(* IEC 61131-3 sources: plcassist-cli/packages/volt-lsp-iec/test-corpus/pro2193/Device/Plc Logic/Application/09 Misc/Library Manager/Standard64, 25 files *)

(* ---- ATOMICREADLINT.fun ---- *)
FUNCTION ATOMICREADLINT : LINT
VAR_INPUT
	PSRC : POINTER TO LINT;
END_VAR
END_FUNCTION

(* ---- ATOMICREADLREAL.fun ---- *)
FUNCTION ATOMICREADLREAL : LREAL
VAR_INPUT
	PSRC : POINTER TO LREAL;
END_VAR
END_FUNCTION

(* ---- ATOMICREADLTIME.fun ---- *)
FUNCTION ATOMICREADLTIME : LTIME
VAR_INPUT
	PSRC : POINTER TO LTIME;
END_VAR
END_FUNCTION

(* ---- ATOMICREADLWORD.fun ---- *)
FUNCTION ATOMICREADLWORD : LWORD
VAR_INPUT
	PSRC : POINTER TO LWORD;
END_VAR
END_FUNCTION

(* ---- ATOMICREADULINT.fun ---- *)
FUNCTION ATOMICREADULINT : ULINT
VAR_INPUT
	PSRC : POINTER TO ULINT;
END_VAR
END_FUNCTION

(* ---- ATOMICWRITELINT.fun ---- *)
FUNCTION ATOMICWRITELINT : BOOL
VAR_INPUT
	PDEST : POINTER TO LINT;
	LIVALUE : LINT;
END_VAR
END_FUNCTION

(* ---- ATOMICWRITELREAL.fun ---- *)
FUNCTION ATOMICWRITELREAL : BOOL
VAR_INPUT
	PDEST : POINTER TO LREAL;
	LRVALUE : LREAL;
END_VAR
END_FUNCTION

(* ---- ATOMICWRITELTIME.fun ---- *)
FUNCTION ATOMICWRITELTIME : BOOL
VAR_INPUT
	PDEST : POINTER TO LTIME;
	LTVALUE : LTIME;
END_VAR
END_FUNCTION

(* ---- ATOMICWRITELWORD.fun ---- *)
FUNCTION ATOMICWRITELWORD : BOOL
VAR_INPUT
	PDEST : POINTER TO LWORD;
	LWVALUE : LWORD;
END_VAR
END_FUNCTION

(* ---- ATOMICWRITEULINT.fun ---- *)
FUNCTION ATOMICWRITEULINT : BOOL
VAR_INPUT
	PDEST : POINTER TO ULINT;
	ULIVALUE : ULINT;
END_VAR
END_FUNCTION

(* ---- WCONCAT.fun ---- *)
FUNCTION WCONCAT : WSTRING(255)
VAR_INPUT
	STR1 : WSTRING(255);
	STR2 : WSTRING(255);
END_VAR
END_FUNCTION

(* ---- WDELETE.fun ---- *)
FUNCTION WDELETE : WSTRING(255)
VAR_INPUT
	STR : WSTRING(255);
	LEN : INT;
	POS : INT;
END_VAR
END_FUNCTION

(* ---- WFIND.fun ---- *)
FUNCTION WFIND : INT
VAR_INPUT
	STR1 : WSTRING(255);
	STR2 : WSTRING(255);
END_VAR
END_FUNCTION

(* ---- WINSERT.fun ---- *)
FUNCTION WINSERT : WSTRING(255)
VAR_INPUT
	STR1 : WSTRING(255);
	STR2 : WSTRING(255);
	POS : INT;
END_VAR
END_FUNCTION

(* ---- WLEFT.fun ---- *)
FUNCTION WLEFT : WSTRING(255)
VAR_INPUT
	STR : WSTRING(255);
	SIZE : INT;
END_VAR
END_FUNCTION

(* ---- WLEN.fun ---- *)
FUNCTION WLEN : INT
VAR_INPUT
	STR : WSTRING(255);
END_VAR
END_FUNCTION

(* ---- WMID.fun ---- *)
FUNCTION WMID : WSTRING(255)
VAR_INPUT
	STR : WSTRING(255);
	LEN : INT;
	POS : INT;
END_VAR
END_FUNCTION

(* ---- WREPLACE.fun ---- *)
FUNCTION WREPLACE : WSTRING(255)
VAR_INPUT
	STR1 : WSTRING(255);
	STR2 : WSTRING(255);
	L : INT;
	P : INT;
END_VAR
END_FUNCTION

(* ---- WRIGHT.fun ---- *)
FUNCTION WRIGHT : WSTRING(255)
VAR_INPUT
	STR : WSTRING(255);
	SIZE : INT;
END_VAR
END_FUNCTION

(* ---- LCTD.fb ---- *)
FUNCTION_BLOCK LCTD
VAR_INPUT
	CD : BOOL;
	LOAD : BOOL;
	PV : LWORD;
END_VAR
VAR_OUTPUT
	Q : BOOL;
	CV : LWORD;
END_VAR
VAR
	M : BOOL;
END_VAR
END_FUNCTION_BLOCK

(* ---- LCTU.fb ---- *)
FUNCTION_BLOCK LCTU
VAR_INPUT
	CU : BOOL;
	RESET : BOOL;
	PV : LWORD;
END_VAR
VAR_OUTPUT
	Q : BOOL;
	CV : LWORD;
END_VAR
VAR
	M : BOOL;
END_VAR
END_FUNCTION_BLOCK

(* ---- LCTUD.fb ---- *)
FUNCTION_BLOCK LCTUD
VAR_INPUT
	CU : BOOL;
	CD : BOOL;
	RESET : BOOL;
	LOAD : BOOL;
	PV : LWORD;
END_VAR
VAR_OUTPUT
	QU : BOOL;
	QD : BOOL;
	CV : LWORD;
END_VAR
VAR
	MU : BOOL;
	MD : BOOL;
	RU : BOOL;
	RD : BOOL;
END_VAR
END_FUNCTION_BLOCK

(* ---- LTOF.fb ---- *)
FUNCTION_BLOCK LTOF
VAR_INPUT
	IN : BOOL;
	PT : LTIME;
END_VAR
VAR_OUTPUT
	Q : BOOL;
	ET : LTIME;
END_VAR
VAR
	M : BOOL;
	STARTTIME : LTIME;
END_VAR
END_FUNCTION_BLOCK

(* ---- LTON.fb ---- *)
FUNCTION_BLOCK LTON
VAR_INPUT
	IN : BOOL;
	PT : LTIME;
END_VAR
VAR_OUTPUT
	Q : BOOL;
	ET : LTIME;
END_VAR
VAR
	M : BOOL;
	STARTTIME : LTIME;
END_VAR
END_FUNCTION_BLOCK

(* ---- LTP.fb ---- *)
FUNCTION_BLOCK LTP
VAR_INPUT
	IN : BOOL;
	PT : LTIME;
END_VAR
VAR_OUTPUT
	Q : BOOL;
	ET : LTIME;
END_VAR
VAR
	STARTTIME : LTIME;
END_VAR
END_FUNCTION_BLOCK
